(* IEC 61131-3 sources: PLC-Static-Analysis/modules/plc-rules/src/test/resources/PLCA-Q007, 2 files *)

(* ---- compliant.st ---- *)
FUNCTION F_Twice : INT
VAR_INPUT
    n : INT;
END_VAR
F_Twice := F_Plus(n, n);
END_FUNCTION

FUNCTION F_Plus : INT
VAR_INPUT
    a : INT;
    b : INT;
END_VAR
F_Plus := a + b;
END_FUNCTION

FUNCTION_BLOCK FB_Timer
METHOD Pulse : BOOL
VAR_INPUT
    bIn : BOOL;
END_VAR
Pulse := THIS^.Pulse(bIn, T#1S);
END_METHOD
METHOD Pulse : BOOL
VAR_INPUT
    bIn : BOOL;
    tLength : TIME;
END_VAR
Pulse := bIn;
END_METHOD
END_FUNCTION_BLOCK

FUNCTION Equal : BOOL
VAR_INPUT
    expected : STRING;
    actual : STRING;
END_VAR
Equal := Equal(expected := TRUE, actual := expected = actual);
END_FUNCTION

(* ---- noncompliant.st ---- *)
FUNCTION F_Rec : INT
VAR_INPUT
    n : INT;
END_VAR
IF n > 0 THEN
    F_Rec := F_Rec(n - 1); // PLCA-Q007
END_IF
END_FUNCTION

FUNCTION F_A : INT
VAR_INPUT
    n : INT;
END_VAR
F_A := F_B(n); // PLCA-Q007
END_FUNCTION

FUNCTION F_B : INT
VAR_INPUT
    n : INT;
END_VAR
F_B := F_A(n);
END_FUNCTION

FUNCTION_BLOCK FB_Tree
METHOD Visit : BOOL
Visit := THIS^.Visit(); // PLCA-Q007
END_METHOD
END_FUNCTION_BLOCK
